PROGRAM MAIN
VAR
	
tempVar		: BOOL;

END_VAR

END_PROGRAM

(* stored: Version 1.1.0.1
   POU MAIN: Id {b4d59aae-968d-46c5-ba60-3ec141f83cb2}, SpecialFunc None *)
